Fanuc KAREL source: kb00116.KL

-- PROVISIONAL review KL for V770-1; original PC SHA256 98483bc4afe6d13691f8effa13337424c7ae7a976065578987208203e333c5e5
-- Incomplete behavior may be omitted. Consult companion uncertainty JSON. Do not deploy.
PROGRAM KB00116
%NOLOCKGROUP
VAR
  P1 : REAL
  RESULT : REAL
BEGIN
  -- UNRESOLVED_PC offsets 5-16; opcodes 2E,23
  -- UNRESOLVED_PC offsets 21-36; opcodes 27,22,76,23
  -- UNRESOLVED_PC offsets 41-45; opcodes 7F
END KB00116
